FUNCTION_BLOCK FB_FastClose
VAR_INPUT
    fStopPos : LREAL;
END_VAR
VAR_OUTPUT
    Closed   : BOOL;;
END_VAR
VAR
    iMotionStage       : I_MotionStage;
    bStarted : BOOL;
END_VAR

IF (iMotionStage = 0)  THEN
    RETURN;
END_IF

Closed := FALSE;
IF 	bStarted THEN
    IF iMotionStage.MotionStatus.bDone THEN
        Closed := TRUE;
        bStarted := FALSE;
    END_IF
END_IF

//FB_Init is always available implicitly and it is used primarily for initialization.
//The return value is not evaluated. For a specific influence, you can also declare the
//methods explicitly and provide additional code there with the standard initialization
//code. You can evaluate the return value.
METHOD FB_Init: BOOL
VAR_INPUT
    bInitRetains: BOOL; // TRUE: the retain variables are initialized (reset warm / reset cold)
    bInCopyCode: BOOL;  // TRUE: the instance will be copied to the copy code afterward (online change)
    iMotionStage : I_MotionStage;
END_VAR
THIS^.iMotionStage := iMotionStage ;
END_METHOD

METHOD Start : BOOL
VAR_INPUT
END_VAR
// Issue move command
iMotionStage.AbsoluteMoveDefault(
   Position     := fStopPos,
   Velocity     := iMotionStage.MotionCmd.fVelocity,
);
bStarted := TRUE;
END_METHOD

END_FUNCTION_BLOCK

(* stored: Version 1.1.0.1
   POU FB_FastClose: Id {0e94abec-494d-4612-9922-721fd3573be3}, SpecialFunc None
   Method FB_Init: Id {690160e3-2846-4668-b6a4-f85d1b586479}
   Method Start: Id {8f6e7839-24ed-4da1-9332-4bca9bff8b25} *)
